(* IEC 61131-3 sources: ICSQuartz/compiler/libs/wrappers/codesys, 1 file *)

(* ---- Common.st ---- *)
/****************************************
Author: Corban Villa
Date: June 16, 2023
Description: This file will wrap the SysFile library
*****************************************/

// https://help.codesys.com/api-content/2/codesys/3.5.14.0/en/_cds_datatype_uxint_xword/
TYPE __XWORD : LWORD;
END_TYPE
